Staubli VAL3: cycle_stop.pgx

public program cycle_stop()
begin
  rs:bToStopCycle=true
  stopMove()
  wait(rs:bIsCycle==false)
  rs:bToStopCycle=false
  logMsg("PLC:stopcycle")
end
